(* IEC 61131-3 sources: kns-pump-station/src/POUs/Time/FB_ScaledClock, 11 files *)

(* ---- FB_ScaledClock.decl.st ---- *)
// Назначение: часы контура с ускорением имитации — источник времени PL.I_TimeSource для
//             устройств, станции, журнала (GVL_Time.fbClockMain) и модели (GVL_Time.fbClockModel).
//             Now() = база + (LTIME() − база_реальная) · k; смена k (Update в начале цикла задачи)
//             перебазирует часы, время монотонно. При k = 1 часы совпадают с LTIME(). Ручной режим
//             (SetManual, AdvanceL) — для интеграционных тестов: время меняется только шагами.
// Автор:      kr0nsch
// Версия:     0.1.0
// Документ:   docs/DESIGN.md, раздел 10; docs/ARCHITECTURE.md, раздел 11
FUNCTION_BLOCK FB_ScaledClock IMPLEMENTS PL.I_TimeSource
VAR
    lrScaleAct   : LREAL := 1.0;     // действующий коэффициент k, 1…SIM_TIME_SCALE_MAX
    ltBaseScaled : LTIME;            // время контура в момент последнего перебазирования
    ltBaseReal   : LTIME;            // LTIME() в тот же момент
    xManual      : BOOL;             // ручной режим: Now() = ltManual
    ltManual     : LTIME := LTIME#1H;   // старт не с нуля (как FB_FakeTime)
    xInit        : BOOL;             // базы заданы первым вызовом Now или Update
END_VAR

(* ---- AdvanceL.method.decl.st ---- *)
// Ручной режим: продвинуть время контура на шаг (вне ручного режима вызов ничего не делает)
METHOD PUBLIC AdvanceL
VAR_INPUT
    ltStep : LTIME;      // шаг
END_VAR

(* ---- AdvanceL.method.impl.st ---- *)
IF xManual THEN
    ltManual := ltManual + ltStep;
END_IF

(* ---- Now.method.decl.st ---- *)
// Время контура, нс; не убывает. В ручном режиме — ltManual
METHOD PUBLIC Now : LTIME
VAR
    ltReal : LTIME;   // системное время этого вызова
END_VAR

(* ---- Now.method.impl.st ---- *)
IF xManual THEN
    Now := ltManual;
    RETURN;
END_IF

ltReal := LTIME();
IF NOT xInit THEN
    // первый вызов: при k = 1 часы совпадают с системным временем
    xInit := TRUE;
    ltBaseReal := ltReal;
    ltBaseScaled := ltReal;
END_IF
Now := ScaledAt(ltReal := ltReal);

(* ---- ScaledAt.method.decl.st ---- *)
// Время контура для системного времени ltReal: ltBaseScaled + (ltReal − ltBaseReal) · k.
// Разность считается только при ltReal > ltBaseReal (LTIME без знака, L7 контракта библиотеки)
METHOD PRIVATE ScaledAt : LTIME
VAR_INPUT
    ltReal : LTIME;      // системное время
END_VAR
VAR
    ltElapsed : LTIME;   // прошло системного времени с перебазирования
END_VAR

(* ---- ScaledAt.method.impl.st ---- *)
IF ltReal <= ltBaseReal THEN
    ScaledAt := ltBaseScaled;
    RETURN;
END_IF

ltElapsed := ltReal - ltBaseReal;
IF lrScaleAct <= 1.0 THEN
    // k = 1 (Update не даёт меньше): без перевода в LREAL — точно при любой длительности
    ScaledAt := ltBaseScaled + ltElapsed;
ELSE
    // LREAL точен до 2^53 нс (≈ 104 сут); дальше округление монотонно
    ScaledAt := ltBaseScaled + ULINT_TO_LTIME(LREAL_TO_ULINT(ULINT_TO_LREAL(LTIME_TO_ULINT(ltElapsed)) * lrScaleAct));
END_IF

(* ---- SetManual.method.decl.st ---- *)
// Ручной режим для интеграционных тестов: xOn = TRUE — Now() = ltStart и дальше меняется только
// AdvanceL. xOn = FALSE — возврат к системному времени: часы продолжают от ручного времени
// (перебазирование), время не идёт назад
METHOD PUBLIC SetManual
VAR_INPUT
    xOn     : BOOL;      // включить ручной режим
    ltStart : LTIME;     // время контура в начале ручного режима (при xOn = TRUE)
END_VAR

(* ---- SetManual.method.impl.st ---- *)
IF xOn THEN
    xManual := TRUE;
    ltManual := ltStart;
ELSIF xManual THEN
    xManual := FALSE;
    xInit := TRUE;
    ltBaseScaled := ltManual;
    ltBaseReal := LTIME();
END_IF

(* ---- Update.method.decl.st ---- *)
// Начало цикла задачи: коэффициент ускорения LIMIT(1, rTimeScale, SIM_TIME_SCALE_MAX), не конечное
// значение → 1. При смене коэффициента — перебазирование: время контура продолжается без скачка
METHOD PUBLIC Update
VAR_INPUT
    rTimeScale : REAL;      // запрошенный коэффициент (GVL_Sim.stSimCfg.rTimeScale или 1)
END_VAR
VAR
    lrScaleNew : LREAL;     // коэффициент после ограничения
    ltReal     : LTIME;     // системное время перебазирования
END_VAR

(* ---- Update.method.impl.st ---- *)
IF PL.F_IsFinite(rIn := rTimeScale) THEN
    lrScaleNew := REAL_TO_LREAL(LIMIT(1.0, rTimeScale, GVL_Const.SIM_TIME_SCALE_MAX));
ELSE
    lrScaleNew := 1.0;
END_IF

ltReal := LTIME();
IF NOT xInit THEN
    xInit := TRUE;
    ltBaseReal := ltReal;
    ltBaseScaled := ltReal;
END_IF

IF lrScaleNew <> lrScaleAct THEN
    // перебазирование одним чтением системного времени: Now() непрерывно в точке смены
    ltBaseScaled := ScaledAt(ltReal := ltReal);
    ltBaseReal := ltReal;
    lrScaleAct := lrScaleNew;
END_IF
